Fanuc KAREL source: kt00034.KL

-- PROVISIONAL review KL for V770-1; original PC SHA256 4fd0593edd455d1562ac70ec86b7b224041847fd7510957fc1b917a05e7ab989
-- Incomplete behavior may be omitted. Consult companion uncertainty JSON. Do not deploy.
PROGRAM KT00034
%NOLOCKGROUP
VAR
  I1 : INTEGER
  I2 : INTEGER
  OUT : REAL
BEGIN
  -- UNRESOLVED_PC offsets 5-16; opcodes 2E,23
  -- UNRESOLVED_PC offsets 21-32; opcodes 2E,23
  -- UNRESOLVED_PC offsets 37-48; opcodes 2E,23
  -- UNRESOLVED_PC offsets 53-64; opcodes 2E,23
  -- UNRESOLVED_PC offsets 69-89; opcodes 21,21,53,64,23
  -- UNRESOLVED_PC offsets 94-98; opcodes 7F
END KT00034
